// Heure UTC en unités de 100 ns depuis 1601 (FILETIME), comme les horodatages échangés avec la HMI
FUNCTION F_NowUtc : LINT

F_NowUtc := ULINT_TO_LINT(F_GetSystemTime());

END_FUNCTION

(* stored: Version 1.1.0.1, ProductVersion 3.1.4024.12
   POU F_NowUtc: Id {e229d065-0d65-50ba-8ee1-2b30720212e2}, SpecialFunc None *)
